// TIA Portal V19 export
// export: Created 2026-10-15T09:44:04.2450986Z, ExportSetting WithDefaults, DisplayName Totally Integrated Automation Portal, DisplayVersion V19, DisplayName TIA Portal Openness, DisplayVersion V19, DisplayName TIA Portal Version Control Interface, DisplayVersion V19, DisplayName STEP 7 Professional, DisplayVersion V19, DisplayName STEP 7 Safety, DisplayVersion V19, DisplayName WinCC Basic/Comfort/Advanced, DisplayVersion V19, DisplayName WinCC Unified, DisplayVersion V19
DATA_BLOCK "ROLL_State"   // DB1
{ S7_Optimized_Access := 'TRUE' }
VERSION : 0.1
// stored: AutoNumber true, DBAccessibleFromOPCUA true, DBAccessibleFromWebserver true, IsOnlyStoredInLoadMemory false, IsRetainMemResEnabled false, IsWriteProtectedInAS false, MemoryReserve 100
   VAR RETAIN
      "M" : Array[0..255, 0..7] of Bool;
      S5Timers { S7_SetPoint := 'True'} : Array[0..127] of "ROLL_TimerState";
      S5Counters { S7_SetPoint := 'True'} : Array[0..127] of "ROLL_CounterState";
      CurrentProgram : Int := 1;
   END_VAR
BEGIN
   "M"[0,4] := TRUE;
END_DATA_BLOCK
